// TIA Portal V21 export
// export: Created 2026-08-21T20:18:50.8353644Z, ExportSetting None, DisplayName Totally Integrated Automation Portal, DisplayVersion V21, DisplayName STEP 7 Professional, DisplayVersion V21, DisplayName STEP 7 Safety, DisplayVersion V21, DisplayName Tech WebApplication, DisplayVersion V21, DisplayName WinCC Basic/Comfort/Advanced, DisplayVersion V21, DisplayName WinCC Professional, DisplayVersion V21, DisplayName WinCC Unified, DisplayVersion V21
FUNCTION "FIT100" : Void   // FC4, FBD
{ S7_Optimized_Access := 'TRUE' }
// stored: SetENOAutomatically false
   VAR_TEMP
      Temp : "DigVal";
      Temp_1 : "DigVal";
   END_VAR
BEGIN

REGION Network 1: MonAnL
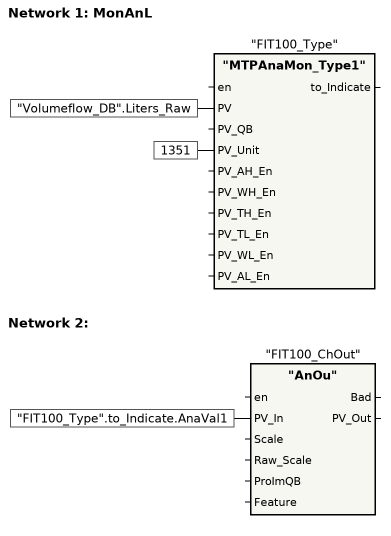
   "FIT100_Type"(PV := "Volumeflow_DB".Liters_Raw, PV_Unit := 1351);   // "MTPAnaMon_Type1"
END_REGION

REGION Network 2
   "FIT100_ChOut"(PV_In := "FIT100_Type".to_Indicate.AnaVal1);   // "AnOu"
END_REGION
END_FUNCTION
